// TIA Portal V21 export
// export: Created 2026-10-23T20:43:17.746482Z, ExportSetting WithDefaults, DisplayName Totally Integrated Automation Portal, DisplayVersion V21 Update 1, DisplayName SINAMICS Startdrive Advanced, DisplayVersion V21 HF2, DisplayName SINAMICS Startdrive G110M, G120, G120C, G120D, G120P, G115D, DisplayVersion V21 HF2, DisplayName SINAMICS Startdrive G130, G150, S120, S150, G200, G220, S200, S210, S220, Innomotics MVD, DisplayVersion V21 HF2, DisplayName STEP 7 Professional, DisplayVersion V21 Update 1, DisplayName STEP 7 Safety, DisplayVersion V21, DisplayName Tech WebApplication, DisplayVersion V21, DisplayName WinCC Basic/Comfort/Advanced, DisplayVersion V21 Update 1, DisplayName WinCC Unified, DisplayVersion V21 Update 1
FUNCTION_BLOCK "FB_AnaDoubleAssign"   // FB13, SCL
TITLE = Analyzer: output assigned twice
{ S7_Optimized_Access := 'TRUE' }
VERSION : 0.1
// Rule C26e: Motor is assigned twice in one cycle
// stored: AutoNumber true, IsIECCheckEnabled false, IsRetainMemResEnabled false, MemoryReserve 100, SetENOAutomatically false, UDAEnableTagReadback false
   VAR_INPUT
      Start : Bool;   // Start
      Stop : Bool;   // Stop
   END_VAR
   VAR_OUTPUT
      Motor : Bool;   // Motor on
   END_VAR
BEGIN

       #Motor := #Start;
       #Motor := #Motor AND NOT #Stop;
END_FUNCTION_BLOCK
